PROGRAM MAIN
VAR
	
END_VAR

RunStudent();

END_PROGRAM

(* stored: Version 1.1.0.1, ProductVersion 3.1.4024.12
   POU MAIN: Id {9ecac31e-5ed6-4cd3-98a5-d9ce44e3a319}, SpecialFunc None *)
